Fanuc KAREL source: ka00014.KL

PROGRAM KA00014
%STACKSIZE=65535
%PRIORITY=65535
%NOLOCKGROUP
VAR
SRC : REAL
DST : REAL
BEGIN
SRC=2.0
DST=SRC
END KA00014
